FUNCTION_BLOCK SK_MoveAxis (* A skill primitive: one action of one piece of equipment (move the axis, run the pump, weigh). It can be called on its own over OPC UA, or be a step of a bigger skill. Inside: SKILL_Core (state machine and OPC UA methods), a parameter block per parameter, SC_ (its contract: what this skill does and when it is done), SKILL_Run (one run, the same for every primitive) and EP_ (the equipment as the skill sees it). Technical: Skill primitive MoveAxis: Head to Position, measured down from the limit switch; the direction follows from where it is (parameters: Position [mm] 0.0..60.0, default 0.0). OPC UA Start(Session, parameters...)/Stop/Abort/Reset(Session) -> [Accepted, ErrorID]; START/HALT/ABORT/RESET from a parent -> SUCCESS or FAILURE(ErrorID) *)
  (* Standard: 61499-2 *)
  (* Version 0.1, 2026-09-28, Project contributors, AAU Smart Production Lab *)
  PACKAGE capping;
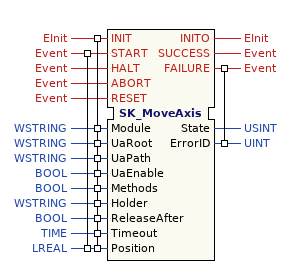
  EVENT_INPUT
    INIT : EInit WITH Module, UaRoot, UaPath, UaEnable, Methods, Holder, ReleaseAfter, Timeout, Position; (* Initialise: its OPC UA nodes and its equipment's channels *)
    START WITH Position; (* Start a run, from the parent (a step of a sequence): no session check *)
    HALT; (* Stop the run, from the parent *)
    ABORT; (* Abort: everything off at once *)
    RESET; (* Reset from Failed or Aborted to Idle *)
  END_EVENT
  EVENT_OUTPUT
    INITO : EInit; (* Initialised: the next block of the INIT chain goes on *)
    SUCCESS; (* The run succeeded (the results are set) *)
    FAILURE WITH ErrorID; (* The run failed (ErrorID) *)
  END_EVENT
  VAR_INPUT
    Module : WSTRING; (* The module's name; its local channels are named after it (loc[<Module>/...]) *)
    UaRoot : WSTRING; (* The module's OPC UA folder, e.g. /Objects/Filling *)
    UaPath : WSTRING; (* This skill's OPC UA folder below UaRoot, e.g. /Skills/Dispensing *)
    UaEnable : BOOL; (* Publish on OPC UA *)
    Methods : BOOL; (* Offer the OPC UA methods Start, Stop, Abort, Reset (FALSE: a step, run by its parent) *)
    Holder : WSTRING; (* The name the equipment is held under: the skill's own, or for a step the skill it belongs to *)
    ReleaseAfter : BOOL := TRUE; (* Give up the equipment when the run ends (FALSE: the next step keeps it) *)
    Timeout : TIME := T#30000ms; (* How long the run may take before it fails with Timeout (3) *)
    Position : LREAL := 0.0; (* Parameter Position mm, 0.0 to 60.0: Where to move to *)
  END_VAR
  VAR_OUTPUT
    State : USINT; (* Skill state: 0 Idle, 1 Running, 2 Stopping, 3 Succeeded, 4 Failed, 5 Aborted *)
    ErrorID : UINT; (* Error code: 0 none, 1 PreconditionViolated, 2 InvariantViolated, 3 Timeout, 4 NotReady, 5 NotPermitted, 6 Busy, 7 Interrupted, 8 OutOfRange *)
  END_VAR
  (* Group SkillControl: State machine and OPC UA: Start(Session, parameters) with the range check, Stop, Abort, Reset; State, parameters and results published *)
  (* Group Execution: What the skill is (its contract) and one run of it, the same for every primitive *)
  (* Group Equipment: The equipment as the skill sees it: its state in, the command out *)
  FBS
    Control : modlib::SKILL_Core; (* The skill's state machine (SKILL_Core): checks a client's Start, publishes State and ErrorID, offers Stop, Abort and Reset over OPC UA, and starts the run when it may begin. *) {SET_ATTRIBUTE(GroupName, SkillControl)}
    Contract : capping::SC_MoveAxis; (* What this skill is (its SC_ type): the command it sends, how long it may run, and when it may start, is done, and must stop. *) {SET_ATTRIBUTE(GroupName, Execution)}
    UaStart : iec61499::net::SERVER_2_2; (* The OPC UA method Start: a client's call arrives here with its session id and the parameters; Control's answer (Accepted, ErrorID) goes back to the client. *) {SET_ATTRIBUTE(GroupName, SkillControl)}
    Par_Position : modlib::SKILL_Param_LREAL(Lower := 0.0, Upper := 60.0); (* The parameter Position: its default, the check of a client's value against its limits, and the value held for the run. *) {SET_ATTRIBUTE(GroupName, SkillControl)}
    PubParams : iec61499::net::PUBLISH_1; (* Writes the parameter values of the current run to OPC UA (Parameters/...). *) {SET_ATTRIBUTE(GroupName, SkillControl)}
    Run : modlib::SKILL_Run; (* One run (SKILL_Run, the same in every primitive): waits for the equipment, checks the contract's precondition, sends the command and watches the conditions until the skill is done. *) {SET_ATTRIBUTE(GroupName, Execution)}
    Port : capping::EP_LinearAxis; (* The equipment as this skill sees it (EP_): its state in (to the contract), the commands from the run (over the adapter AEquipment). *) {SET_ATTRIBUTE(GroupName, Equipment)}
  END_FBS
  EVENT_CONNECTIONS
    Control.START_RSP TO UaStart.RSP;
    UaStart.IND TO Par_Position.CHECK;
    Control.RUN TO Par_Position.LATCH;
    Par_Position.CHECKED TO Control.START_REQ;
    Par_Position.LATCHED TO PubParams.REQ;
    PubParams.INITO TO PubParams.REQ;
    INIT TO Control.INIT;
    Control.INITO TO Contract.INIT;
    Contract.INITO TO UaStart.INIT;
    UaStart.INITO TO Par_Position.INIT;
    Par_Position.INITO TO PubParams.INIT;
    PubParams.INITO TO Run.INIT;
    Run.INITO TO Port.INIT;
    Port.INITO TO INITO;
    START TO Control.START;
    HALT TO Control.HALT;
    ABORT TO Control.ABORT;
    RESET TO Control.RESET;
    Control.SUCCESS TO SUCCESS;
    Control.FAILURE TO FAILURE;
    Par_Position.LATCHED TO Contract.START;
    Control.HALT_SEQ TO Run.HALT;
    Control.ABORT_SEQ TO Run.ABORT;
    Control.RUN_STOPPING TO Control.STOPPING_DONE;
    Run.DONE TO Control.EXECUTE_DONE;
    Run.FAILED TO Control.EXECUTE_FAILED;
    Run.HALTED TO Control.EXECUTE_FAILED;
    Port.STATE TO Contract.SAMPLE;
  END_CONNECTIONS
  DATA_CONNECTIONS
    Control.StartMethodId TO UaStart.ID;
    UaStart.RD_1 TO Control.Session;
    Control.Accepted TO UaStart.SD_1;
    Control.StartError TO UaStart.SD_2;
    UaStart.RD_2 TO Par_Position.Requested;
    Control.CalledByClient TO Par_Position.CalledByClient;
    Par_Position.Value TO PubParams.SD_1;
    Par_Position.AllInRange TO Control.ParamsInRange;
    Module TO Control.Module;
    UaRoot TO Control.UaRoot;
    UaPath TO Control.UaPath;
    UaEnable TO Control.UaEnable;
    Methods TO Control.Methods;
    Methods TO UaStart.QI;
    Control.State TO State;
    Control.ErrorID TO ErrorID;
    UaRoot TO Contract.UaRoot;
    UaPath TO Contract.UaPath;
    Timeout TO Contract.Timeout;
    UaEnable TO PubParams.QI;
    Contract.IdParams TO PubParams.ID;
    Position TO Par_Position.Default;
    Par_Position.Value TO Contract.Position;
    Holder TO Run.Holder;
    ReleaseAfter TO Run.ReleaseAfter;
    Run.ErrorID TO Control.ExecuteError;
    Module TO Port.Module;
    Port.ActualPosition TO Contract.ActualPosition;
    Port.Homed TO Contract.Homed;
    Port.Moving TO Contract.Moving;
    Port.EqHolder TO Contract.EqHolder;
    Run.EquipmentFree TO Control.EquipmentFree;
  END_CONNECTIONS
  ADAPTER_CONNECTIONS
    Contract.Run TO Run.Contract;
    Run.Equipment TO Port.Skill;
  END_CONNECTIONS
END_FUNCTION_BLOCK
